// TIA Portal V20 export
// export: Created 2026-10-20T12:39:36.0649577Z, ExportSetting WithDefaults, DisplayName Totally Integrated Automation Portal, DisplayVersion V20 Update 6, DisplayName TIA Portal Openness, DisplayVersion V20 Update 6, DisplayName TIA Portal Version Control Interface, DisplayVersion V20 Update 6, DisplayName SINAMICS Startdrive Advanced, DisplayVersion V20 SP1, DisplayName SINAMICS Startdrive G130, G150, S120, S150, SINAMICS MV, G220, S200, S210, DisplayVersion V20 SP1, DisplayName SINAMICS Startdrive G110M, G120, G120C, G120D, G120P, G115D, DisplayVersion V20 SP1, DisplayName STEP 7 Professional, DisplayVersion V20 Update 6, DisplayName STEP 7 Safety, DisplayVersion V20 Update 2, DisplayName WinCC Basic/Comfort/Advanced, DisplayVersion V20 Update 6, DisplayName WinCC Unified, DisplayVersion V20 Update 6
DATA_BLOCK "Control_DB"   // DB69
{ S7_Optimized_Access := 'TRUE' }
VERSION : 0.1
// stored: AutoNumber true, DBAccessibleFromOPCUA true, IsOnlyStoredInLoadMemory false, IsRetainMemResEnabled false, IsWriteProtectedInAS false, MemoryReserve 100
   VAR
      ECnv_Sys { S7_SetPoint := 'True'} : Array[1..5] of "ECnv_Control";
      LCnv_Sys { S7_SetPoint := 'True'} : Array[1..5] of "Cnv_VTD_Control";
      VTD_Sys { S7_SetPoint := 'True'} : Array[1..5] of "VTD_Control";
      WCS_OPC_Control { S7_SetPoint := 'True'} : Array[1..5] of "WMS_OPC_UA";
      Shuttles_Position : Array[1..23] of Struct
         x : DInt;
         y : DInt;
         Charging : Bool;
      END_STRUCT;
      VTDBarcode_Station : Array[1..5] of "Barcode_Station_UDT";
      Pallet_ID_Received : Array[1..3] of Bool;
      Gate_Station : Array[1..12] of "Gate_Station_UDT";
   END_VAR
BEGIN
   LCnv_Sys[4].Cnv_Level[1..8].Cnv2.Safety_Stop_Cnrl.Inputs.DP_Extended := TRUE;
   LCnv_Sys[5].Cnv_Level[1..8].Cnv2.Safety_Stop_Cnrl.Inputs.DP_Extended := TRUE;
END_DATA_BLOCK
